{attribute 'pack_mode' := '1'}
TYPE S_TURBINEDATA :
STRUCT
	WindSpeed			: REAL;
	WindDirection		: REAL;
	PowerGen			: REAL;
	YawAng				: REAL;
	RotorSpeed			: REAL;
	PitchAngle			: REAL;
	PitchAngleSpt		: REAL;
	GenTorque			: REAL;
END_STRUCT
END_TYPE

(* stored: Version 1.1.0.1
   DUT S_TURBINEDATA: Id {1e57f15f-ebcc-4899-8f91-5fae8db087cd} *)
